TYPE E_CamMachineState :
(
    CAM_STATE_DISABLED := 0,
    CAM_STATE_POWERING,
    CAM_STATE_IDLE,
    CAM_STATE_REFERENCING_MASTER,
    CAM_STATE_REFERENCING_SLAVE,
    CAM_STATE_BUILDING_TABLE,
    CAM_STATE_LOADING_TABLE,
    CAM_STATE_READY,
    CAM_STATE_CAMMING_IN,
    CAM_STATE_STARTING_MASTER,
    CAM_STATE_RUNNING,
    CAM_STATE_STOPPING_MASTER,
    CAM_STATE_RELEASING_STOP,
    CAM_STATE_CAMMING_OUT,
    CAM_STATE_RETURNING_SLAVE,
    CAM_STATE_RESETTING,
    CAM_STATE_FAULT
);
END_TYPE

(* stored: Version 1.1.0.1, ProductVersion 3.1.4024.16
   DUT E_CamMachineState: Id {a621df35-176a-4f38-be79-d4f1f9f312a9} *)
